FUNCTION_BLOCK GenericBistableDeviceModel (* Migrated from IEC 61131-3 ST *)
  (* Standard: 61499-2 *)
  (* Version 1.0, 2026-11-06, st2fb *)
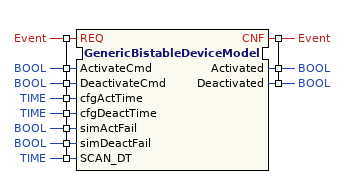
  EVENT_INPUT
    REQ WITH ActivateCmd, DeactivateCmd, cfgActTime, cfgDeactTime, simActFail, simDeactFail, SCAN_DT;
  END_EVENT
  EVENT_OUTPUT
    CNF WITH Activated, Deactivated;
  END_EVENT
  VAR_INPUT
    ActivateCmd : BOOL;
    DeactivateCmd : BOOL;
    cfgActTime : TIME := T#1s;
    cfgDeactTime : TIME := T#1s;
    simActFail : BOOL;
    simDeactFail : BOOL;
    SCAN_DT : TIME;
  END_VAR
  VAR_OUTPUT
    Activated : BOOL;
    Deactivated : BOOL;
  END_VAR
  VAR
    TransitionDelay_IN : BOOL;
    TransitionDelay_PT : TIME;
    TransitionDelay_Q : BOOL;
    TransitionDelay_ET : TIME;
    TransitionDelay_STATE : INT;
    TransitionDelay_PREV_IN : BOOL;
    TransitionDelay_START_TIME : TIME;
    ST2FB_NOW : TIME;
    vState : INT := 0;
    vStateOld : INT := 3;
  END_VAR
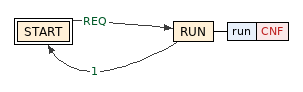
  EC_STATES
    START;
    RUN : run -> CNF;
  END_STATES
  EC_TRANSITIONS
    START TO RUN := REQ;
    RUN TO START := 1;
  END_TRANSITIONS
  ALGORITHM run IN ST:
ST2FB_NOW := ST2FB_NOW + SCAN_DT;
CASE vState OF
  0:
    IF vState <> vStateOld THEN
      TransitionDelay_IN := FALSE;
      IF (TransitionDelay_STATE = 0) AND NOT TransitionDelay_PREV_IN AND TransitionDelay_IN THEN
        TransitionDelay_STATE := 1;
        TransitionDelay_Q := FALSE;
        TransitionDelay_START_TIME := ST2FB_NOW;
      ELSE
        IF NOT TransitionDelay_IN THEN
          TransitionDelay_ET := T#0s;
          TransitionDelay_Q := FALSE;
          TransitionDelay_STATE := 0;
        ELSIF TransitionDelay_STATE = 1 THEN
          IF TransitionDelay_START_TIME + TransitionDelay_PT <= ST2FB_NOW THEN
            TransitionDelay_STATE := 2;
            TransitionDelay_Q := TRUE;
            TransitionDelay_ET := TransitionDelay_PT;
          ELSE
            TransitionDelay_ET := ST2FB_NOW - TransitionDelay_START_TIME;
          END_IF;
        END_IF;
      END_IF;
      TransitionDelay_PREV_IN := TransitionDelay_IN;
      vStateOld := vState;
    END_IF;
    TransitionDelay_IN := ActivateCmd AND NOT simActFail;
    TransitionDelay_PT := cfgActTime;
    IF (TransitionDelay_STATE = 0) AND NOT TransitionDelay_PREV_IN AND TransitionDelay_IN THEN
      TransitionDelay_STATE := 1;
      TransitionDelay_Q := FALSE;
      TransitionDelay_START_TIME := ST2FB_NOW;
    ELSE
      IF NOT TransitionDelay_IN THEN
        TransitionDelay_ET := T#0s;
        TransitionDelay_Q := FALSE;
        TransitionDelay_STATE := 0;
      ELSIF TransitionDelay_STATE = 1 THEN
        IF TransitionDelay_START_TIME + TransitionDelay_PT <= ST2FB_NOW THEN
          TransitionDelay_STATE := 2;
          TransitionDelay_Q := TRUE;
          TransitionDelay_ET := TransitionDelay_PT;
        ELSE
          TransitionDelay_ET := ST2FB_NOW - TransitionDelay_START_TIME;
        END_IF;
      END_IF;
    END_IF;
    TransitionDelay_PREV_IN := TransitionDelay_IN;
    IF TransitionDelay_Q THEN
      vState := 1;
    END_IF;
  1:
    IF vState <> vStateOld THEN
      TransitionDelay_IN := FALSE;
      IF (TransitionDelay_STATE = 0) AND NOT TransitionDelay_PREV_IN AND TransitionDelay_IN THEN
        TransitionDelay_STATE := 1;
        TransitionDelay_Q := FALSE;
        TransitionDelay_START_TIME := ST2FB_NOW;
      ELSE
        IF NOT TransitionDelay_IN THEN
          TransitionDelay_ET := T#0s;
          TransitionDelay_Q := FALSE;
          TransitionDelay_STATE := 0;
        ELSIF TransitionDelay_STATE = 1 THEN
          IF TransitionDelay_START_TIME + TransitionDelay_PT <= ST2FB_NOW THEN
            TransitionDelay_STATE := 2;
            TransitionDelay_Q := TRUE;
            TransitionDelay_ET := TransitionDelay_PT;
          ELSE
            TransitionDelay_ET := ST2FB_NOW - TransitionDelay_START_TIME;
          END_IF;
        END_IF;
      END_IF;
      TransitionDelay_PREV_IN := TransitionDelay_IN;
      vStateOld := vState;
    END_IF;
    TransitionDelay_IN := DeactivateCmd AND NOT simDeactFail;
    TransitionDelay_PT := cfgDeactTime;
    IF (TransitionDelay_STATE = 0) AND NOT TransitionDelay_PREV_IN AND TransitionDelay_IN THEN
      TransitionDelay_STATE := 1;
      TransitionDelay_Q := FALSE;
      TransitionDelay_START_TIME := ST2FB_NOW;
    ELSE
      IF NOT TransitionDelay_IN THEN
        TransitionDelay_ET := T#0s;
        TransitionDelay_Q := FALSE;
        TransitionDelay_STATE := 0;
      ELSIF TransitionDelay_STATE = 1 THEN
        IF TransitionDelay_START_TIME + TransitionDelay_PT <= ST2FB_NOW THEN
          TransitionDelay_STATE := 2;
          TransitionDelay_Q := TRUE;
          TransitionDelay_ET := TransitionDelay_PT;
        ELSE
          TransitionDelay_ET := ST2FB_NOW - TransitionDelay_START_TIME;
        END_IF;
      END_IF;
    END_IF;
    TransitionDelay_PREV_IN := TransitionDelay_IN;
    IF TransitionDelay_Q THEN
      vState := 0;
    END_IF;
END_CASE;
Activated := vState = 1;
Deactivated := vState = 0;
  END_ALGORITHM
END_FUNCTION_BLOCK
